FUNCTION_BLOCK FB_Gr01Angle
(*

The function block used to control axis .

Constructor: 		Patryk Panylo
Company:		E. Riexinger GmbH
Date:			28.04.2015
Version:			1.00

Date:			Revision:		Who:				Comment
dd.mm.yyyy		x.xx			Initials			comment

*)
VAR_INPUT
	(* Input variables / Eingang Variablen *)
	(* --- Axis / Achse --- *)
	bEnable						:BOOL;						(* Axis present *)
	bOccupied					:BOOL;						(* Axis is occupied *)

	(* --- Machine state / Maschinenzustand --- *)
	etMachineMode				:ET_MachineMode;			(* Machine mode *)
	etMachineState				:ET_MachineState;			(* Machine state *)
	bMachineStandstill			:BOOL;						(* Machine standstill *)

	(* --- Safety & releases / Sicherheit & Freigaben --- *)
	bNoEStop					:BOOL;						(* No ermergency Stop / Keine Notaus *)
	bPowerSupplyOn				:BOOL;						(* Power supply on / Leitung eingeschaltet *)
	bSafetyOK					:BOOL;						(* Safety ok / Sicherheit i.o *)
	bSafetyDriveEnabled			:BOOL;						(* Safety drive enable *)
	bCtrlInterrupt				:BOOL;						(* Control interrupt *)
	bMoveRelease				:BOOL;						(* Move release *)
	bMoveInterrupt				:BOOL;						(* Move Interrupt *)
	bPlusRelease				:BOOL;						(* Plus move release *)
	bMinusRelease				:BOOL;						(* Minus move release *)

	(* --- Limits / Endlagen --- *)
	bHWSignalLimitMax			:BOOL;						(* Signal position limit switch maximum *)
	bHWSignalLimitMin			:BOOL;						(* Signal position limit switch minimum *)
	lrSoftLimitMax				:LREAL;						(* Position limit switch maximum *)
	lrSoftLimitMin				:LREAL;						(* Position limit switch minimum *)

	(* --- Commands / Befehle --- *)
	bExeReset					:BOOL;						(* Execute auto reset *)
	bExeHome					:BOOL;						(* Execute home *)
	bExeMoveAbs					:BOOL;						(* Execute move absolut *)
	bExeMoveVelo				:BOOL;						(* Execute move velo *)
	bExeGearIn					:BOOL;						(* Execute gear in *)
	bExeGearOut					:BOOL;						(* Execute gear out *)
	bExeStop					:BOOL;						(* Execute move stop *)
	bConfirmAlarm				:BOOL;						(* Confirm alarm *)

	(* --- Manual mode / Handbetrieb --- *)
	bTipPlus					:BOOL;						(* Manual tip in plus direction *)
	bTipMinus					:BOOL;						(* Manual tip in minus direction *)
	lrManualVelocity			:LREAL;						(* Value of velocity in manual motion [mm/s] *)

	(* --- Motion parameters / Bewegungsparameter --- *)
	lrTargetPosition			:LREAL;						(* Absolute target position *)
	lrAutoVelocity				:LREAL;						(* Value of velocity in auto motion [mm/s] *)
	lrVelocityNoRef				:LREAL;						(* Velocity if has no reference [mm/s] *)
	bVelocityLimitEn			:BOOL;						(* Enable velocity limit *)
	lrVelocityMin				:LREAL;						(* Velocity minimum [%] *)
	lrVelocityMax				:LREAL;						(* Velocity maximum [%] *)
	lrAcceleration				:LREAL;						(* Value of the acceleration (always positive) *)
	lrDeceleration				:LREAL;						(* Value of deceleration (always positive) *)
	lrJerk						:LREAL;						(* Value of jerk (always positive) *)

	(* --- Override --- *)
	lrOverride					:LREAL;						(* Override *)
	bExtOverrideEn				:BOOL;						(* External override enable *)
	lrExtOverride				:LREAL;						(* External override *)

	(* --- Gearing / Getriebe --- *)
	dnRatioNumerator			:DINT;						(* Gear ratio numerator. Alternatively, the gear ratio can be specified in the numerator as a floating comma value, if the denominator is 1. *)
	udnRatioDenominator			:UDINT;						(* Gear ratio denominator *)

	(* --- Drive / Antrieb --- *)
	snModesOfOperation			:SINT;						(* Modes of drive operation *)
	bEngineTorqueLimitEn		:BOOL;						(* Enable engine torque limit *)
	lrEngineTorque				:LREAL;						(* Engine torque [%] *)
	bPosLagMonitoringEn			:BOOL;						(* Enable position lag monitoring *)
	tControllerOff				:TIME := T#60S;				(* Time to switch controller off *)

	(* --- Scaling & encoder / Skalierung & Geber --- *)
	lrScalingNum				:LREAL := 1.0;				(* Effective distance per rev. Numerator [technical units] *)
	udnScalingDenom				:UDINT := 1;				(* Effective distance per rev. Denominator [INC] *)
	bWithAbsoluteEncoder		:BOOL;						(* Encoder is an absolute one / Absolutwertgeber *)
	udnIncEnc					:UDINT;						(* Value of encoder increment *)
	lrOriginShift				:LREAL;						(* Origin shift position *)

	(* --- System --- *)
	lrTaskCycle					:LREAL := 0.002;			(* Cycle time of the task [sec], 0.002[s] => 2ms *)
	tAdsTimeOut					:TIME := T#2S;				(* Timout for ads commands *)
END_VAR
VAR_OUTPUT
	(* Output variables / Ausgang Variablen *)
	(* --- Status --- *)
	bCtrlEnabled				:BOOL;						(* Controller enabled *)
	bNotMoving					:BOOL;						(* Axis not moving *)
	bStandStill					:BOOL;						(* Added by Dustin for 633_Hilton) Axis stands stil*)
	bReferenced					:BOOL;						(* Axis referenced *)
	bCoupled					:BOOL;						(* Axis coupled *)

	(* --- Actual values / Istwerte --- *)
	lrActPosition				:LREAL;						(* Actual position [mm] *)
	lrActAbsPosition			:LREAL;						(* Actual absolut position [mm] *)
	lrActVelocity				:LREAL;						(* Actual velocity [mm/s] *)
	lrVeloMax					:LREAL;						(* Velocity limit maximum *)

	(* --- Limits / Endlagen --- *)
	bHardLimitMaxExceeded		:BOOL;						(* Position limit switch maximum is exceeded *)
	bHardLimitMinExceeded		:BOOL;						(* Position limit switch minimum is exceeded *)
	bSoftLimitMaxExceeded		:BOOL;						(* Position limit switch maximum is exceeded *)
	bSoftLimitMinExceeded		:BOOL;						(* Position limit switch minimum is exceeded *)

	(* --- Safety / Sicherheit --- *)
	bSafetyLock					:BOOL;						(* Safety lock*)
	bSafetyDriveEnable			:BOOL;						(* Safety drive enable *)

	(* --- Errors / Fehler --- *)
	bErrorTerminal				:BOOL;						(* Error Axis terminal *)
	bErrorCtrlEnabled			:BOOL;						(* Error Axis controller enabled *)
	
END_VAR
VAR_IN_OUT	
	(* Input Output variables / Ausgang Variablen *)
	bHomeCompleted				:BOOL;						(* Home completed *)
	Drive						:ST_STOEBERSI6SC6CIA402_REF;
	Axis						:AXIS_REF;
	MasterAxis					:AXIS_REF;
END_VAR
VAR
	(* Enummerations *)

	(* Variables *)
	sAdsAddr					:STRING(23);					(* AmsNetId of the EtherCAT master device.*)
	unSlaveAddr					:UINT;							(* Address of the slave device.*)

	nTorqueLimitMax				:INT := 100;					(* The torque limit (absolute value). Value range in %: -200 ... 200 ... 200 *)

	lrVeloLimitMax				:LREAL;
	lrVeloLimitMin				:LREAL;

	sTerminalStatus				:STRING;

	(* References *)

	(* Interfaces *)

	(* Instances *)
	fbTerminalDiagnosis			:FB_TerminalDiagnosis;
	rtMachineStandstill			:R_TRIG;
	tonAxisEnabled				:TON;

	fbController				:FB_STOEBER_AxisController;
	fbMoveManual				:FB_STOEBER_AxisMoveManual;
	fbMoveAuto					:FB_STOEBER_AxisMoveAuto;
	(*fbDriveLink				:FB_STOEBER_DriveLink;*)
	fbForce						:FB_ScalingOffset;
	fbForceCtrl					:FB_ForceController;
	fbCoolingOff				:FB_SignalHandlingDelay;
END_VAR


IF NOT bEnable								(* Signal FB enable *)
THEN

	RETURN;
END_IF

(* Old Axis Ref from Tc2) 
(* ControllerConfig *)
stControllerConfig.lrKp := 0.018;						(* Tuning parameter, proportional gain *)
stControllerConfig.lrTi := 0.0;							(* Tuning parameter, time of integral *)
stControllerConfig.lrTd := 0.0;						(* Tuning parameter, time of differential *)
stControllerConfig.lrPreCtrlVelo := 0.01; 				(* Feedforward velocity precontrol wieghting =  0..1 *)
stControllerConfig.lrVeloKpFilter := 1.0;				(* Velocity filter - proportional gain *)
stControllerConfig.tVeloT1Filter := t#100ms;			(* Velocity filter - time constant *)
stControllerConfig.tDeadTime  := t#100ms;				(* Dead time *)
stControllerConfig.lrDeltaMax := 10.0;					(* Maximum difference between two actual position values filtered [inc] *)
stControllerConfig.lrVeloMin := -7.8; 					(* Velocity limit minimum [deg / sec] *)
stControllerConfig.lrVeloMax  := 7.8; 					(* Velocity limit maximum [deg / sec] *)
stControllerConfig.lrDeadZone := 10.0;					(* Dead zone *)

(* Encoder configuration *)
stEncoderConfig.dwModuloValue := 8192; 			(* Maximum encoder modulo value e.g 1048576 [inc] *)
stEncoderConfig.etScalingMethod := ET_ScalingMethod_eSMLinear;

(* Interface *)
stAxis.stScaling.dwModuloValue := 8192; 		(* Maximum encoder modulo value 4294967295 dword *)
stAxis.stAxisCtrl.bEnable := Axis.stPlcToNc.stBaseDevice.bEnable;
stAxis.stAxisStates.bOperational := Axis.stNcToPlc.stBaseDevice.bEnabled;
stAxis.stScaling.etScalingMethod := ET_ScalingMethod_eSMLinear;
stAxis.stScaling.lrTaskCycle := lrTaskCycle;
stAxis.stScaling.udnScalingDenom := udnScalingDenom; (* inc *)
stAxis.stScaling.lrScalingNum := lrScalingNum; (* deg *)
stAxis.stScaling.lrScaleFactor := udnScalingDenom / lrScalingNum;
stAxis.stPosition.lrOffsetPos := lrOriginShift;
stAxis.stLimitSwitches.lrSWPosLimitMin := lrSoftLimitMin;
stAxis.stLimitSwitches.lrSWPosLimitMax := lrSoftLimitMax;

A_AxisLink();
A_AxisGetStatus();
A_AxisController();
A_AxisMoveManual();
A_AxisMoveAuto();
A_AxisTerminalDiag();
A_AxisAlarm();


lrSpeedFactor := F_kAngleActuatorSpeedLin(
						bEnable := TRUE,
						lrActAngle := lrActPosition,
						lrAngleOffset := 56.6,  (* [deg] *)
						lrMultiplier := 0.755,
						lrOffset := 0.24
					);

Axis.stPlcToNc.stBaseDevice.stFastRefereneValue.nSpeed := LREAL_TO_INT(INT_TO_LREAL(Axis.stPlcToNc.stBaseDevice.stFastRefereneValue.nSpeed) * lrSpeedFactor);

*)

ACTION A_AxisAlarm:

(* Axis errors *)
tonAxisEnabled(
	IN := fbController.bEnable
		AND fbController.bRegulatorOn
		AND NOT fbController.bStatusDelay,
	PT := fbController.tStatusDelay + t#2s
);

bErrorCtrlEnabled := tonAxisEnabled.Q;
END_ACTION

ACTION A_AxisController:

(* Axis controller *)
fbController(
    bEnable := TRUE,
	etMachineMode := etMachineMode,
	etMachineState := etMachineState,
	bNoEStop := bNoEStop,
	bRegulatorOn := bNoEStop
				      AND bPowerSupplyOn
				      AND bSafetyOk
				      AND SEL(bNotMoving, NOT bCtrlInterrupt, TRUE)
				      AND NOT fbMoveManual.bControllerOff
				      AND NOT fbMoveAuto.bControllerOff,
	bReset := bConfirmAlarm,
	bTerminalOK := fbTerminalDiagnosis.bTerminalOK,
	bExeReset := bExeReset,
	bExeSetPos := FALSE,
	lrSetPosition := lrTargetPosition,
	bExeGearIn := bExeGearIn,
	bExeGearOut := bExeGearOut,
	dnRatioNumerator := dnRatioNumerator,
	udnRatioDenominator := udnRatioDenominator,
	lrOverride := SEL(bExtOverrideEn,
					lrOverride,
					lrOverride*lrExtOverride/100.0),
	bWithAbsoluteEncoder := bWithAbsoluteEncoder,
	bPosLagMonitoringEn := bPosLagMonitoringEn,
	lrPositionBias := 0.0,
	lrSoftLimitMax := lrSoftLimitMax,
	lrSoftLimitMin := lrSoftLimitMin,
	bSignalHWLimitMax:= bHWSignalLimitMax,
	bSignalHWLimitMin := bHWSignalLimitMin,
	lrAcceleration := lrAcceleration,
	lrDeceleration := lrDeceleration,
	lrJerk := lrJerk,
	pDrive := ADR(Drive),
	Axis := Axis,
	MasterAxis := MasterAxis,
	bStatusDelay => bCtrlEnabled,
	lrActPos => lrActPosition,
	lrActAbsPos => lrActAbsPosition,
	lrActVelo => lrActVelocity,
	bNotMoving => bNotMoving,
	bStandStill => bStandStill,
	bReferenced => bReferenced,
	bCoupled => bCoupled,
	lrVeloLimitMax => lrVeloMax,
	bHardLimitMaxExceeded => bHardLimitMaxExceeded,
	bHardLimitMinExceeded => bHardLimitMinExceeded,
	bSoftLimitMaxExceeded => bSoftLimitMaxExceeded,
	bSoftLimitMinExceeded => bSoftLimitMinExceeded
);

bSafetyDriveEnable := fbMoveManual.bSafetyCtrlEnable 
				 	  OR fbMoveAuto.bSafetyCtrlEnable;



(* from Tc2)

(* Axis controller *)
fbController(
    	bEnable := TRUE,
	etMachineMode := etMachineMode,
	etMachineState := etMachineState,
	bRegulatorOn := bNoEStop
				      AND bPowerSupplyOn
				      AND bSafetyOK
                 		      	      AND NOT bCtrlInterrupt
				      AND NOT fbMoveManual.bControllerOff
				      AND NOT fbMoveAuto.bControllerOff,
	bReset := bConfirmAlarm,
	bTerminalOK := fbTerminalDiagnosis.bTerminalOK,
	bExeReset := bExeReset,
	dwRawMotorEncoder := udnIncEnc,
	lrOverride := SEL(bExtOverrideEn,
					lrOverride,
					lrOverride*lrExtOverride/100.0),
	lrEngineTorque := SEL(
						bEngineTorqueLimitEn,
						nTorqueLimitMax,
						(lrEngineTorque) / 1),
	bWithAbsoluteEncoder := bWithAbsoluteEncoder,
	bHWSignalLimitMax := bHWSignalLimitMax,
	bHWSignalLimitMin := bHWSignalLimitMin,
	lrSoftLimitMax := lrSoftLimitMax,
	lrSoftLimitMin := lrSoftLimitMin,
	stEncoderConfig := stEncoderConfig,
	pAxis := ADR(stAxis),
	Axis := Axis,
	bStatusDelay => bCtrlEnabled,
	lrActPos=> ,
	lrActVelo => lrActVelocity,
	bNotMoving => bNotMoving,
	bReferenced => bReferenced,
	bHardLimitMaxExceeded => bHardLimitMaxExceeded,
	bHardLimitMinExceeded => bHardLimitMinExceeded,
	bSoftLimitMaxExceeded => bSoftLimitMaxExceeded,
	bSoftLimitMinExceeded => bSoftLimitMinExceeded
);

lrActPosition := F_LRealRound(fbController.lrActPos,1);
*)
END_ACTION

ACTION A_AxisGetStatus:

(* Get axis status *)
Axis.ReadStatus();
END_ACTION

ACTION A_AxisLink:

(* Get terminal status *)
sAdsAddr := F_CreateAmsNetId(Drive.stTerminalState.stAdsAddr.netId);
unSlaveAddr := Drive.stTerminalState.stAdsAddr.port;
Axis.DriveAddress.NetID := F_CreateAmsNetId(Drive.stTerminalState.stAdsAddr.netId);
Axis.DriveAddress.SlaveAddress := Drive.stTerminalState.stAdsAddr.port;

(* Set drive parameter *)
Drive.stPlcToStoeber.snA541ModesOfOperation := snModesOfOperation;

(*Drive.PlcToStoeber.nA558TargetTorque := SEL(bEngineTorqueLimitEn,
				    nTorqueLimitMax,
				    LREAL_TO_INT(lrEngineTorque / 1.0))*)
END_ACTION

ACTION A_AxisMoveAuto:

(* Move axis auto *)
rtMachineStandstill(CLK := bMachineStandstill);

lrVeloLimitMin := SEL(bVelocityLimitEn, -1 * lrVeloMax, lrVelocityMin);
lrVeloLimitMax := SEL(bVelocityLimitEn, lrVeloMax, lrVelocityMax);


fbMoveAuto(
	bEnable := bNoEStop
			   AND bPowerSupplyOn
			   AND bSafetyOK,
	bOccupied := bOccupied,
	bSafetyCtrlEnabled := bSafetyDriveEnabled,
	bCtrlEnabled := bCtrlEnabled
				      AND bMoveRelease,
	etMachineMode := etMachineMode,
	etMachineState := etMachineState,
	bReset := bConfirmAlarm,
	bCtrlEnable := bCtrlEnabled,
	bExeHome := bExeHome,
	bExeMoveAbs := bExeMoveAbs,
	bExeMoveVelo := bExeMoveVelo,
	bExeStop := bExeStop
			    OR rtMachineStandstill.Q,
	lrPosition := lrTargetPosition,
	lrVelocity := LIMIT(lrVeloLimitMin, lrAutoVelocity, lrVeloLimitMax),
	lrAcceleration := lrAcceleration,
	lrDeceleration := lrDeceleration,
	lrJerk := lrJerk,
	tControllerOff := tControllerOff,
	pDrive := ADR(Drive),
	bHomeCompleted := bHomeCompleted,
	Axis := Axis,
	MasterAxis := MasterAxis
 );
(* From Tc3) 

fbMoveAuto(
	bEnable := bNoEStop
               		    AND bPowerSupplyOn
               		    AND bSafetyOK,
	bCtrlEnabled := bCtrlEnabled
                    		   AND bMoveRelease,
	etMachineMode := etMachineMode,
	etMachineState := etMachineState,
	bReset := bConfirmAlarm,
	bExeHome := bExeHome,
	bExeMoveAbs := bExeMoveAbs,
	bExeMoveVelo := bExeMoveVelo,
	bExeStop := bExeStop
			      OR rtMachineStandstill.Q,
	lrPosition := lrTargetPosition,
	lrVelocity := LIMIT(lrVeloLimitMin, lrAutoVelocity, lrVeloLimitMax),
	lrAcceleration := lrAcceleration,
	lrDeceleration := lrDeceleration,
	lrJerk := lrJerk,
	tControllerOff := tControllerOff,
	stControllerConfig := stControllerConfig,
	pAxis := ADR(stAxis),
	bHomeCompleted := bHomeCompleted,
	Axis := Axis
 );
 
 *)
END_ACTION

ACTION A_AxisMoveManual:

(* Move axis manual *)
fbMoveManual(
	bEnable := bNoEStop
               		    AND bPowerSupplyOn
               		    AND bSafetyOK,
	bCtrlEnabled := bCtrlEnabled
               			    AND bMoveRelease,
	etMachineMode := etMachineMode,
	etMachineState := etMachineState,
	bReset := bConfirmAlarm,
	bMovePlus := bTipPlus,
	bMoveMinus := bTipMinus,
	bLimitMax := bHardLimitMaxExceeded
			       OR bSoftLimitMaxExceeded,
	bLimitMin := bHardLimitMinExceeded
			      OR bSoftLimitMinExceeded,
	bPlusRelease := bPlusRelease,
	bMinusRelease := bMinusRelease,
	lrVelocity := SEL(NOT bReferenced, lrManualVelocity, lrVelocityNoRef),
	tControllerOff := tControllerOff,
	bHomeCompleted := bHomeCompleted,
	Axis := Axis,
	MasterAxis 				:= GVL_Gr00Interface.iAxisDummy,
);

bSafetyLock := fbMoveManual.bMovePlus
                		OR fbMoveManual.bMoveMinus;
END_ACTION

ACTION A_AxisTerminalDiag:

(*Axis terminal diagnosis *)
fbTerminalDiagnosis(
	stTerminalState := Drive.stTerminalState,
	sTerminalStatus => sTerminalStatus
);

bErrorTerminal := NOT fbTerminalDiagnosis.bTerminalOK;
END_ACTION

END_FUNCTION_BLOCK

(* stored: Version 1.1.0.1, ProductVersion 3.1.4024.15
   POU FB_Gr01Angle: Id {55356d1b-1b2b-4ec3-9464-e4dce6e77525}, SpecialFunc None
   Action A_AxisAlarm: Id {64cefd6f-6bba-4c72-a96d-bc952e00de0b}
   Action A_AxisController: Id {cd705a5b-95b6-4c6b-b77f-d7fda30432c2}
   Action A_AxisGetStatus: Id {407ebed2-432b-449e-87bc-1349d7b19c57}
   Action A_AxisLink: Id {17b267a5-3daf-42cc-aef1-ad1a7d1a108c}
   Action A_AxisMoveAuto: Id {ecb8cc8c-5caf-4778-b2b8-51d55fb57cac}
   Action A_AxisMoveManual: Id {d121ea87-82c5-4a44-9e9a-9dbd906b351e}
   Action A_AxisTerminalDiag: Id {39933bb9-04fb-4401-aaae-96fb36b33781} *)
